Fanuc KAREL source: NC0066.KL

-- PROVISIONAL review KL for V940-1; original PC SHA256 24ac9b305348f69286334de9e712197caf62ba846f88e8a3accdb24c0b0eb176
-- Incomplete behavior may be omitted. Consult companion uncertainty JSON. Do not deploy.
PROGRAM NC0066
%NOLOCKGROUP
-- UNRESOLVED_LOCAL_POOL 9 cells at code offset 3; source declarations unknown
-- DIRECT_LOCAL_WORD_ACCESS alone does not prove INTEGER, REAL, or BOOLEAN
BEGIN
  -- V9_EXPOSED_INDEXED_TABLE_HINT layout=0001; 16 counted words exposed once; source arms/runtime held
  -- V9_FOOTER_20_HINT 8 numerical footer links; VM transfer unproved
  -- UNRESOLVED_PC offsets 0-8; opcodes 2B,2C,7B
  -- UNRESOLVED_PC offsets 13-20; opcodes 9D,23
  -- UNRESOLVED_PC offsets 25-54; opcodes 9D,23,9E,2E,22,7A
  -- UNRESOLVED_PC offsets 59-88; opcodes 9D,23,9E,2E,22,7A
  -- UNRESOLVED_PC offsets 93-122; opcodes 9D,23,9E,2E,22,7A
  -- UNRESOLVED_PC offsets 127-156; opcodes 9D,23,9E,2E,22,7A
  -- UNRESOLVED_PC offsets 161-190; opcodes 9D,23,9E,2E,22,7A
  -- UNRESOLVED_PC offsets 195-224; opcodes 9D,23,9E,2E,22,7A
  -- UNRESOLVED_PC offsets 229-258; opcodes 9D,23,9E,2E,22,7A
  -- UNRESOLVED_PC offsets 263-292; opcodes 9D,23,9E,2E,22,7A
  -- UNRESOLVED_PC offsets 297-311; opcodes 21,9D,52,23
  -- UNRESOLVED_PC offsets 316-331; opcodes 20,2C,23
  -- UNRESOLVED_PC offsets 336-351; opcodes 20,2C,23
  -- UNRESOLVED_PC offsets 356-371; opcodes 20,2C,23
  -- UNRESOLVED_PC offsets 376-391; opcodes 20,2C,23
  -- UNRESOLVED_PC offsets 396-411; opcodes 20,2C,23
  -- UNRESOLVED_PC offsets 416-431; opcodes 20,2C,23
  -- UNRESOLVED_PC offsets 436-451; opcodes 20,2C,23
  -- UNRESOLVED_PC offsets 456-471; opcodes 20,2C,23
  -- UNRESOLVED_PC offsets 476-480; opcodes 7F
  -- UNRESOLVED_PC offsets 485-489; opcodes 27,AA
  -- UNRESOLVED_PC offsets 494-498; opcodes 7F
END NC0066
